FUNCTION F_CheckSyntaxString : BOOL (* TRUE if STR does not contain capital letters *)
VAR_INPUT
	str 		:T_MaxString;
	flag 		:T_MaxString;
	sep 		:T_MaxString := '=';
	sufix		:POINTER TO STRING; 					
END_VAR
VAR
	L			:INT;
	prefix1		:T_MaxString;
	prefix2		:T_MaxString;
	
END_VAR


prefix1 := CONCAT(flag, sep);
L := LEN(prefix1);
prefix2 := MID(str, L, 1);

F_CheckSyntaxString := FALSE;

IF LEN(str) > L
THEN
	sufix^ := DELETE(str, L, 1);
	IF prefix1 = prefix2
	THEN
		F_CheckSyntaxString := TRUE;
	END_IF;
END_IF

END_FUNCTION

(* stored: Version 1.1.0.1, ProductVersion 3.1.4024.15
   POU F_CheckSyntaxString: Id {40870304-d26b-46df-8114-6e062cf1568b}, SpecialFunc None *)
